(* IEC 61131-3 sources: sis-interlock-demo/src/POUs/Generated/FB_SisApp, 1 file *)

(* ---- FB_SisApp.decl.st ---- *)
// AUTO-GENERATED by cemgen 1.0.0 — не редактировать: правьте матрицу и запустите
//   python -m cemgen generate <файл матрицы .csv или .xlsx>
// Матрица: SIS-V101-CEM, объект V-101, ревизия B от 2026-10-19, SHA-256 сетки df2ed4841a9453ca
// Назначение: привязка ПАЗ объекта V-101 к образу ввода-вывода: токи 4–20 мА → инж. ед. и
//             достоверность по NE 43, дискретные входы и контроль линии → группы голосования по
//             причинам; вызов FB_SisUnit с конфигурацией GVL_SisCfg; разрешения следствий → выходы
//             xQ*.
// Автор:      kr0nsch; код — генератор cemgen
// Версия:     1.0.0
// Документ:   docs/DESIGN.md, раздел «10. Генератор cemgen»; docs/cause_effect_matrix.md
// ВНИМАНИЕ:   код демонстрационный и не предназначен для систем безопасности. Реальная ПАЗ требует
//             определения SIL, сертифицированных аппаратных и программных средств и валидации по
//             ГОСТ Р МЭК 61511.
FUNCTION_BLOCK FB_SisApp
VAR_INPUT
    itfTime : PL.I_TimeSource;      // 0 — системное время
    itfLog  : I_SisEventSink;       // 0 — без журнала
END_VAR
VAR_IN_OUT
    stIo  : ST_SisIo;               // входы читает, выходы xQ* пишет
    stCmd : ST_SisCmd;              // команды HMI
END_VAR
VAR_OUTPUT
    xTripped   : BOOL := TRUE;                                          // сработало хотя бы одно следствие
    stCemSts   : ST_CauseEffectSts;                                     // состояние матрицы
    astVoteSts : ARRAY[1..GVL_Const.SIS_CAUSES_MAX] OF ST_VotingSts;   // состояние групп голосования
END_VAR
VAR
    fbUnit : FB_SisUnit;                                                // общий узел ПАЗ
    astIn  : ARRAY[1..GVL_Const.SIS_CAUSES_MAX] OF ST_VoteIn;       // входы групп по причинам
END_VAR
